PROGRAM ladderLabel
VAR
	coil: BOOL;
END_VAR

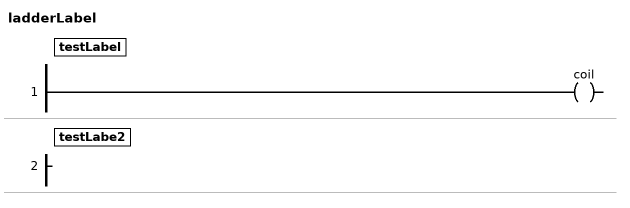
// NETWORK 1
testLabel:
coil := TRUE;

// NETWORK 2
testLabe2: ;

END_PROGRAM

(* stored: Version 1.1.0.1, ProductVersion 3.1.4024.16
   POU ladderLabel: Id {1bd00e36-8301-4b53-a0d5-dff6189ade52}, SpecialFunc None *)
